INTERFACE I_Resettable EXTENDS __SYSTEM.IQueryInterface

METHOD Reset
END_METHOD

END_INTERFACE

(* stored: Version 1.1.0.1
   Itf I_Resettable: Id {19d8f4e6-7b9d-4ea2-919b-db452d7c134c}
   Method Reset: Id {8def40b3-3d7b-4e44-9e8b-d4bea9900221} *)
